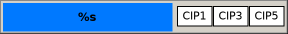
VISUALIZATION vis_FB_Element_CIP  // 288x34
VAR_IN_OUT
	fb: FB_Element;
END_VAR
    Rectangle (0,0 288x34)
    Textfield (2,2 171x30), "%s", text variable: fb.sElementID
    RoundedRectangle (177,6 35x20), "CIP1"
        tap fb.bTakePosInCIPBuffer_Partial
    RoundedRectangle (213,6 35x20), "CIP3"
        tap fb.bTakePosInCIPBuffer_Detergent
    RoundedRectangle (249,6 35x20), "CIP5"
        tap fb.bTakePosInCIPBuffer_Full
END_VISUALIZATION

(* stored: Version 1.1.0.1, ProductVersion 3.1.4024.12
   Visu vis_FB_Element_CIP: Id {dcaa9652-771c-4e66-a1b6-53630db990b2} *)
